(* CODESYS project cognex_insight.library
   DefaultNamespace: KOSTAL.AF2024.Drivers.Camera.Cognex_InSight
   DocFormat: reStructuredText
   Description: Provides communication via TcpIp or Ethernet/IP to Cognex InSight cameras.
   Author: Frank Dümpelmann, Martí Puig (F2R Automation)
   Title: KOSTAL.AF2024.Drivers.Camera.Cognex_InSight
   Version: 3.0.0.0
   Company: KOSTAL GmbH & Co.KG
   Placeholder: KOSTAL.AF2024.Drivers.Camera.Cognex_InSight

Project tree, tasks and I/O mapping:
  libraries: KOSTAL.AF2024.Core.ListOf, 1.0.0.0 (KOSTAL GmbH & Co.KG); KOSTAL.AF2024.Core.Process, 1.1.0.0 (KOSTAL GmbH & Co.KG); KOSTAL.AF2024.Core.Settings, 1.0.0.0 (KOSTAL GmbH & Co.KG); KOSTAL.AF2024.Core.StringTools, 1.0.0.0 (KOSTAL GmbH & Co.KG); KOSTAL.AF2024.Core.System, 1.0.0.0 (KOSTAL GmbH & Co.KG); KOSTAL.AF2024.Drivers.Camera.I_Camera, 2.0.0.0 (KOSTAL GmbH & Co.KG); Tc2_Standard, 3.4.5.0 (Beckhoff Automation GmbH); Tc2_System, 3.9.1.0 (Beckhoff Automation GmbH); Tc2_TcpIp, 3.4.2.0 (Beckhoff Automation GmbH); Tc2_Utilities, 3.9.2.0 (Beckhoff Automation GmbH)
  EthernetIP/
    DUT/
      Result/
        interface I_T_Result_Base: Clear, ResultArray
      data type _E_THIS_EIP
      data type _T_InspectionResult
      data type ST_IN_EIP
      data type ST_OUT_EIP
    function block FB_InSight_EIP [ST]: _a0_StepFail, _a0_StepInit, _a1_finish, _a1_idle, _a2_callTrigger, _a2_changeProgNum, _a2_inspection_Result, _connectControl, _FBmain, _resetfault, Ex_SetProgramNumber, Ex_Trigger, Ex_Trigger_ProgramNumber, FaultReset, LinkResult, Fault, ProgNo, ResultPass, State, FBmain
    interface I_InSight_EIP: Fault
  Project Information/
    function F_GetCompany [ST]
    function F_GetTitle [ST]
    function F_GetVersion [ST]
  TcpIp/
    DUT/
      Info/
        interface I_T_Info_TcpIp: ApplicationVersion, CopyTo, DateOfBuild, MacAddress, MonitorVersion, SerialNumber
        interface I_T_Info_TcpIp_CopyFrom: CopyFrom
        interface I_T_Info_TcpIp_Owner: ApplicationVersion, Clear, CopyFrom, DateOfBuild, MacAddress, MonitorVersion, SerialNumber
        function block T_Info_TcpIp [ST]: ApplicationVersion, Clear, CopyFrom, CopyTo, DateOfBuild, MacAddress, MonitorVersion, SerialNumber
      Internal/
        data type _E_PrgType_TcpIp
        data type _E_THIS_TcpIp
      data type E_BuilderVersion_TcpIp
      data type E_Command_TcpIp
      data type E_ProgLocation_TcpIp
    function block FB_InSight_Explorer_TcpIp [ST]: FB_init, _c1_Receive, _c1_Send, _c1_Socket, _connectionInit, _catchMacId, _catchPrgId, _catchPrgName, _foundEtx, _isCommandAccept, _isPasswordRequest, _isUserAccrepted, _isUserRequest, _isWelcome, _SplitData, _getCommand, _a3_GetData, _a3_GetData_DS, _a3_GetData_ETH, _a0_stepFail, _a0_stepInit, _a1_failure, _a1_Finish, _a1_Idle, _a2_Login, _a3_GetInfo, _a3_GetPrgId, _a3_GetPrgName, _a3_SetOffline, _a3_SetOnline, _a3_SetReqPrgById, _a3_SetReqPrgByName, _a3_Trigger, _FBmain, Ex_GetInfo, Ex_GetProgamNumber, Ex_GetProgramName, Ex_SetProgramName, Ex_SetProgramNumber, Ex_Trigger, Ex_Trigger_ProgName, Ex_Trigger_ProgramNumber, CommandPort, CommandTimeOut, IP, Data, DigitalSignalRuntime, DisableComplexResult, Info, ProgLocation, ResultPass, State, FBmain
    function block FB_InSight_VisionSuite_TcpIp [ST]: _catchMacId, _getCommand, SheetName
    interface I_InSight_TcpIp: Ex_GetInfo, Ex_GetProgamNumber, Ex_GetProgramName, Ex_SetProgramName, Ex_Trigger_ProgName, CommandPort, CommandTimeOut, IP, Data, DigitalSignalRuntime, DisableComplexResult, Info, ProgLocation
  Version/
    global variables Global_Version
*)

// EthernetIP/DUT/_E_THIS_EIP
{attribute 'qualified_only'}
{attribute 'strict'}
TYPE INTERNAL _E_THIS_EIP :
(
	idle	:= 0,
	trig,			
	trigPrgNum,
	chgprgnum	
) UINT;
END_TYPE

// EthernetIP/DUT/_T_InspectionResult
TYPE INTERNAL _T_InspectionResult : ARRAY[1..480] OF BYTE; END_TYPE

// EthernetIP/DUT/ST_IN_EIP
{attribute 'pack_mode' := '0'} 
TYPE ST_IN_EIP :
	STRUCT	
		TriggerReady 					: BIT;		//0.0
		TriggerACK						: BIT;		//0.1
		noName_0_0						: BIT;		//0.2
		MissedAcq							: BIT;		//0.3
		OfflineReason_1				: BIT;		//0.4		
		OfflineReason_2				: BIT;		//0.5
		OfflineReason_3				: BIT;		//0.6
		Online								: BIT;		//0.7
		SystemBusy						: BIT;		//1.0
		InspectionCompleted		: BIT;      //1.1
		ResultsBufferOverrun	: BIT;      //1.2
		ResultsValid					: BIT;      //1.3
		CommandExecuting			: BIT;      //1.4
		CommandComplete				: BIT;      //1.5
		CommandFailed					: BIT;      //1.6
		Error									: BIT;      //1.7
		SetUserDataAck				: BIT;		//2.0
		noName_1_0						: BIT;      //2.1
		noName_1_1						: BIT;      //2.2
		ExposureComplete			: BIT;      //2.3
		JobPass								: BIT;      //2.4
		TestRunReady					: BIT;      //2.5
		noName_2_0						: BIT;      //2.6
		noName_2_1						: BIT;      //2.7
		SoftEventACK_0				: BIT;		//3.0
		SoftEventACK_1				: BIT;      //3.1
		SoftEventACK_2				: BIT;      //3.2
		SoftEventACK_3				: BIT;      //3.3
		SoftEventACK_4				: BIT;      //3.4
		SoftEventACK_5				: BIT;      //3.5
		SoftEventACK_6				: BIT;      //3.6
		SoftEventACK_7				: BIT;      //3.7
		ErrorCode							: INT;
		noName_3_0						: BYTE;
		noName_3_1						: BYTE;
		CurrentJobID					: UINT;		
		AcquisitionID					: UINT;
		IspectionID						: UINT;
		InspectionResultCode	: INT;
		InspectionResult			: _T_InspectionResult;
	END_STRUCT
END_TYPE

// EthernetIP/DUT/ST_OUT_EIP
{attribute 'pack_mode' := '0'} 
TYPE ST_OUT_EIP :
	STRUCT
		TriggerEnable					: BIT; 		//0.0								
		Trigger								: BIT; 	    //0.1
		BufferResultsEnable		: BIT; 	    //0.2
		InspectionResultsACK	: BIT; 	    //0.3
		ExecuteCommand				: BIT; 	    //0.4
		noName_0_0						: BIT; 	    //0.5
		noName_0_1						: BIT; 	    //0.6
		SetOffline						: BIT; 	    //0.7
		noName_1							: BYTE;		//1
		SetUserData						: BIT; 		//2.0
		noName_2_0						: BIT; 	    //2.1
		ClearError						: BIT; 	    //2.2
		ClearExposureComplete	: BIT; 	    //2.3
		noName_3_0						: BIT; 	    //2.4
		noName_3_1						: BIT;      //2.5
		noName_3_2						: BIT; 	    //2.6
		noName_3_3						: BIT;      //2.7
		SoftEvent_0						: BIT; 		//3.0
		SoftEvent_1						: BIT;      //3.1
		SoftEvent_2						: BIT;      //3.2
		SoftEvent_3						: BIT;      //3.3
		SoftEvent_4						: BIT;      //3.4
		SoftEvent_5						: BIT;      //3.5
		SoftEvent_6						: BIT;      //3.6
		SoftEvent_7						: BIT;      //3.7
		CommandID							: UINT;	
		noName_4_0						: BYTE; 	
		noName_4_1						: BYTE; 	
		UserData							: _T_InspectionResult;// ARRAY[0..487] OF BYTE; 
	END_STRUCT
END_TYPE

// TcpIp/DUT/Internal/_E_PrgType_TcpIp
{attribute 'qualified_only'}
{attribute 'strict'}
TYPE INTERNAL _E_PrgType_TcpIp :
(
	Number := 0,
	Name
) UINT;
END_TYPE

// TcpIp/DUT/Internal/_E_THIS_TcpIp
{attribute 'qualified_only'}
{attribute 'strict'}
TYPE INTERNAL _E_THIS_TcpIp :
(
	Idle := 0,
	GetInfo,

	Trigger,
	TriggerPrgNo,
	TriggerPrgName,

	SetOnline,
	GetOnline,

	SetProgramId,
	GetProgramId,

	SetProgramName,
	GetProgramName,

	ReadVersion,
	ReadOperationMode
) UINT;
END_TYPE

// TcpIp/DUT/E_BuilderVersion_TcpIp
{attribute 'qualified_only'}
{attribute 'strict'}
TYPE E_BuilderVersion_TcpIp :
(
	InSightExplorer 	:= 0,
	InSigtVisionSuite	:= 1
);
END_TYPE

// TcpIp/DUT/E_Command_TcpIp
{attribute 'qualified_only'}
{attribute 'strict'}
TYPE E_Command_TcpIp :
(
	GetInfo := 0,
	UserName,
	Password,
	SetOnline,
	SetOffline,
	GetOnline,
	GetPrgId,
	SetPrgId,
	GetPrgName,
	SetPrgName,
	Trigger,
	GetFormatstring
);
END_TYPE

// TcpIp/DUT/E_ProgLocation_TcpIp
{attribute 'qualified_only'}
{attribute 'strict'}
TYPE E_ProgLocation_TcpIp :
(
	None := 0,
	FlashMemory,
	RamDisk,
	SD_Card
);
END_TYPE

// Version/Global_Version
{attribute 'TcGenerated'}
{attribute 'no-analysis'}
{attribute 'linkalways'}
// This function has been automatically generated from the project information.
VAR_GLOBAL CONSTANT
	{attribute 'const_non_replaced'}
	stLibVersion_KOSTAL_AF2024_Drivers_Camera_Cognex_InSight : ST_LibVersion := (iMajor := 3, iMinor := 0, iBuild := 0, iRevision := 0, nFlags := 0, sVersion := '3.0.0.0');
END_VAR

// EthernetIP/DUT/Result/I_T_Result_Base
INTERFACE PUBLIC I_T_Result_Base EXTENDS KOSTAL_AF2024_Core_System.I_Interface

METHOD PUBLIC Clear
VAR

END_VAR
END_METHOD

PROPERTY PUBLIC ResultArray : REFERENCE TO _T_InspectionResult
GET
END_GET
END_PROPERTY

END_INTERFACE

// EthernetIP/FB_InSight_EIP
FUNCTION_BLOCK FB_InSight_EIP IMPLEMENTS I_InSight_EIP//, _I_T_Result

VAR
	{region 'EthernetIP Communications'}
		ECatState			AT %I*	: UINT;	//link to EtherCat State from {Device x (ECAT EIP Scanner (EL6652))}.Inputs.State
		InSightState	AT %I*	: UINT;	//link to {InSight 2000 Series}.Inputs.State
	
		InSight_IN 	AT %I*	: ST_IN_EIP; //link with Continious mode ATTENTION be sure, that the Array-Nodes are collapsed
		InSight_OUT AT %Q*	: ST_OUT_EIP; //link with Continious mode ATTENTION be sure, that the Array-Nodes are collapsed
															
//		InSight_IN	: POINTER TO ST_IN_EIP;
//		InSight_OUT	: POINTER TO ST_OUT_EIP;
	{endregion}
                            	                     	
	_step	: KOSTAL_AF2024_Core_Process.FB_processStep_Flow;	//Use the “_Flow” step to save runtime. 

	_THIS_CALLED			: _E_THIS_EIP;
	_THIS_IN_PROCESS	: _E_THIS_EIP;

	_state	: KOSTAL_AF2024_Core_Process.T_plcState;
	
	{region 'Functionality'}
		//Inputs 
		_Reset	: BOOL;
		_prgNum	: UINT;
															
		//Outputs               	
		_InspectionOK				: BOOL;
		//_InspectionNOK			: BOOL;
		//_refResult	: REFERENCE TO _T_InspectionResult;
		_Iresult	: I_T_Result_Base;	 
 
	{endregion}

	{region 'Static'}
		TON_Change_Job : Tc2_Standard.TON;
	{endregion}
		 

	
		 
	
END_VAR

VAR CONSTANT
	_ADDRESS_Idle						: INT:= 0;
	_ADDRESS_TriggerPrgNum	: INT:= 100;	//Job ID
	_ADDRESS_SetPrgNum			: INT:= 200;	//Job ID
END_VAR

METHOD PROTECTED _a0_StepFail
VAR_INPUT
END_VAR

_state.clear();
_state.fail:= TRUE;
_state.description:= Tc2_Standard.WCONCAT(INT_TO_WSTRING(_step.actual), ". Step does not exist");
END_METHOD

METHOD PROTECTED _a0_StepInit
VAR_INPUT
END_VAR

IF (_THIS_CALLED <> _THIS_IN_PROCESS) AND_THEN (_step.actual <> _ADDRESS_Idle) THEN	_step.init();	END_IF
END_METHOD

METHOD PROTECTED _a1_finish 
VAR_INPUT
END_VAR

_state.clear();

_state.finish := TRUE;
_state.pass:= TRUE;
END_METHOD

METHOD PROTECTED _a1_idle

//Idle process - Clear information from other processes
IF _step.toggle THEN

	InSight_OUT.Trigger								:= FALSE;
	InSight_OUT.TriggerEnable					:= FALSE;
	InSight_OUT.InspectionResultsACK := FALSE;

END_IF


_state.clear();

IF _THIS_CALLED = _E_THIS_EIP.idle THEN

	_THIS_IN_PROCESS:= _THIS_CALLED;

	_state.ready := TRUE;

	
ELSIF _THIS_CALLED = _E_THIS_EIP.chgprgnum THEN

	_THIS_IN_PROCESS:= _THIS_CALLED;

	_state.busy := TRUE;

	_step.set(_ADDRESS_SetPrgNum);
	
	
ELSIF _THIS_CALLED = _E_THIS_EIP.trigPrgNum THEN

	_THIS_IN_PROCESS:= _THIS_CALLED;

	_state.busy := TRUE;

	_InspectionOK:= FALSE;
	
	_step.set(_ADDRESS_TriggerPrgNum);

	
ELSIF _THIS_CALLED = _E_THIS_EIP.trig THEN

	_THIS_IN_PROCESS:= _THIS_CALLED;

	_state.busy := TRUE;

	_InspectionOK:= FALSE;

	_step.set(_ADDRESS_TriggerPrgNum);
	
ELSE

	_THIS_IN_PROCESS:= _E_THIS_EIP.idle;

	_state.finish	:= TRUE;
	_state.fail		:= TRUE;
	_state.description:= 	"Process with this enumeration does not exist!"; 

END_IF
END_METHOD

METHOD PROTECTED _a2_callTrigger
VAR_INPUT
END_VAR

VAR_INST	
	_SubStep		: KOSTAL_AF2024_Core_Process.FB_processStep_Flow;
	_PF_InspectionCompleted	:BOOL;
END_VAR

IF _step.toggle THEN	
	_subStep.init();
	IF _Iresult <> 0 THEN
		_Iresult.Clear();
END_IF	
END_IF

_state.description:= "Method _a2_callTrigger() is running ...";

InSight_OUT.InspectionResultsACK := FALSE;

_subStep.Header();

IF _SubStep.isActive(0) THEN IF InSight_IN.ResultsValid THEN InSight_OUT.InspectionResultsACK := TRUE; ELSE _SubStep.INC(); END_IF END_IF
	
IF _SubStep.isActive(1) THEN IF NOT  InSight_IN.ResultsValid THEN InSight_OUT.TriggerEnable := TRUE ; InSight_OUT.InspectionResultsACK := FALSE; _SubStep.INC(); END_IF END_IF

IF _SubStep.isActive(2) THEN IF  InSight_IN.TriggerReady (*AND NOT _pIN^.InspectionCompleted*) THEN InSight_OUT.Trigger:= TRUE; _SubStep.INC(); END_IF END_IF

IF _SubStep.isActive(3) THEN IF InSight_IN.InspectionCompleted <> _PF_InspectionCompleted THEN InSight_OUT.Trigger := FALSE; _step.INC(); END_IF END_IF

_PF_InspectionCompleted := InSight_IN.InspectionCompleted;
END_METHOD

METHOD PROTECTED _a2_changeProgNum
VAR_INPUT
END_VAR
IF _step.toggle THEN	;	END_IF

_state.description:= "Method _a2_changeProgNum() is running ...";

IF InSight_IN.CurrentJobID > 0 AND InSight_IN.CurrentJobID = _prgNum THEN
	
	InSight_OUT.SetOffline := FALSE;
	TON_Change_Job(IN:= FALSE);

	_step.INC();

ELSE

	InSight_OUT.CommandID := _prgNum;
	InSight_OUT.SetOffline := TRUE;

	IF  NOT InSight_IN.Online AND InSight_IN.OfflineReason_1 THEN
		//TON_Change_Job.PT := T#100MS;
		//TON_Change_Job.IN := TRUE;
		TON_Change_Job(IN:= TRUE, PT:= T#100MS, Q=> , ET=> );
	END_IF

END_IF

InSight_OUT.ExecuteCommand := TON_Change_Job.Q;
END_METHOD

METHOD PROTECTED _a2_inspection_Result
VAR_INPUT
END_VAR

IF _step.toggle THEN	;	END_IF

_state.description:= "Method _a2_inspection_Result() is running ...";

InSight_OUT.TriggerEnable 	:= FALSE ;
_InspectionOK  				:= FALSE;


IF _Iresult <> 0 AND_THEN __ISVALIDREF(_Iresult.ResultArray) THEN
	_Iresult.ResultArray := InSight_IN.InspectionResult;
END_IF


_InspectionOK := InSight_IN.InspectionResult[1] = 1;

_step.INC();
END_METHOD

METHOD PROTECTED _connectControl : BOOL
VAR_INPUT
END_VAR

 
IF ECatState <> 0  THEN

	_connectControl:= FALSE;

	_state.clear();
	_state.fail:= TRUE;
	_state.description:= Tc2_Standard.WCONCAT(UINT_TO_WSTRING(ECatState), ";Error from EtherCAT (EIP-Scanner)");


	_step.init();

ELSIF InSightState <> 0 THEN

	_connectControl:= FALSE;

	_state.clear();
	_state.fail:= TRUE;
	_state.description:= Tc2_Standard.WCONCAT(UINT_TO_WSTRING(InSightState), ";Error from Ethernet IP Connection");

	_step.init();

ELSE
	
	_connectControl:= TRUE;

END_IF
END_METHOD

METHOD PROTECTED _FBmain
VAR_INPUT
END_VAR
// is set duriing FB_Init() method
//_pIN:= ADR(InSight2000_IN[2]);
//_pOUT:= ADR(InSight2000_OUT[2]);


IF NOT _connectControl() THEN RETURN;	END_IF

_a0_StepInit();

_step.Header();

IF _step.isActive(_ADDRESS_Idle) THEN _a1_idle();	END_IF


//Trigger and TriggerPrgNum uses the same steps
IF _step.isActive(_ADDRESS_TriggerPrgNum)			THEN _step.INC();							END_IF
IF _step.isActive(_ADDRESS_TriggerPrgNum + 1)	THEN _a2_changeProgNum();			END_IF
IF _step.isActive(_ADDRESS_TriggerPrgNum + 2)	THEN _a2_callTrigger();				END_IF
IF _step.isActive(_ADDRESS_TriggerPrgNum + 3)	THEN _a2_inspection_Result();	END_IF
IF _step.isActive(_ADDRESS_TriggerPrgNum + 4)	THEN _a1_finish();						END_IF


IF _step.isActive(_ADDRESS_SetPrgNum)			THEN _step.INC();					END_IF
IF _step.isActive(_ADDRESS_SetPrgNum + 1)	THEN _a2_changeProgNum();	END_IF
IF _step.isActive(_ADDRESS_SetPrgNum + 2)	THEN _a1_finish();				END_IF


IF _step.NotFound() THEN _a0_StepFail();	END_IF

_resetfault();
END_METHOD

METHOD PROTECTED _resetfault
VAR_INPUT
END_VAR

IF _Reset AND InSight_IN.Error THEN	InSight_OUT.ClearError := TRUE;
ELSE														InSight_OUT.ClearError := FALSE;
END_IF

_Reset:= FALSE;
END_METHOD

METHOD PUBLIC Ex_SetProgramNumber : BOOL;
VAR_INPUT
	ProgramNumber : UINT;
END_VAR
IF _THIS_CALLED = _E_THIS_EIP.idle THEN //Another process is running: don't start this process!

	_prgNum := ProgramNumber;
	
	_THIS_CALLED := _E_THIS_EIP.chgprgnum;
	
	_FBmain();	//Call sequence via _FBmain
	
	Ex_SetProgramNumber := _THIS_CALLED = _THIS_IN_PROCESS;	//Return true when process was started
	
END_IF
END_METHOD

METHOD Ex_Trigger : BOOL

IF _THIS_CALLED = _E_THIS_EIP.idle THEN //Another process is running: don't start this process!

	_THIS_CALLED := _E_THIS_EIP.trig;
	
	_FBmain();	//Call sequence via _FBmain
	
	Ex_Trigger := _THIS_CALLED = _THIS_IN_PROCESS;	//Return true when process was started

END_IF
END_METHOD

METHOD PUBLIC Ex_Trigger_ProgramNumber : BOOL;
VAR_INPUT
	ProgramNumber : UINT;
END_VAR
IF _THIS_CALLED = _E_THIS_EIP.idle THEN //Another process is running: don't start this process!

	IF ProgramNumber <> 0 THEN	_prgNum := ProgramNumber;	END_IF
	
	_THIS_CALLED := _E_THIS_EIP.trigPrgNum;
	
	_FBmain();	//Call sequence via _FBmain
	
	Ex_Trigger_ProgramNumber := _THIS_CALLED = _THIS_IN_PROCESS;	//Return true when process was started

END_IF
END_METHOD

METHOD PUBLIC FaultReset

_Reset := TRUE;
END_METHOD

METHOD PUBLIC LinkResult
VAR_INPUT
	result 	: I_T_Result_Base;
END_VAR
IF result <> 0 THEN
 _Iresult := result; 
END_IF;
END_METHOD

PROPERTY Fault : bool
GET
Fault := InSight_IN.Error;
END_GET
END_PROPERTY

PROPERTY ProgNo : UINT
GET

ProgNo:=  InSight_IN.CurrentJobID;;
END_GET
END_PROPERTY

PROPERTY ResultPass : BOOL
GET

ResultPass:= _InspectionOK;
END_GET
END_PROPERTY

PROPERTY State : KOSTAL_AF2024_Core_Process.I_T_plcState
GET
State := _state;
END_GET
END_PROPERTY

METHOD FBmain
VAR_INPUT
END_VAR

VAR

END_VAR

IF _THIS_CALLED = _E_THIS_EIP.idle THEN
	_FBmain();
END_IF
_THIS_CALLED:= _E_THIS_EIP.idle;
END_METHOD

END_FUNCTION_BLOCK

// EthernetIP/I_InSight_EIP
INTERFACE I_InSight_EIP EXTENDS KOSTAL_AF2024_Drivers_Camera_I_Camera.I_Camera

PROPERTY Fault : bool
GET
END_GET
END_PROPERTY

END_INTERFACE

// Project Information/F_GetCompany
// This function has been automatically generated from the project information.
{attribute 'signature_flag' := '1073741824'}
{attribute 'TcGenerated'}
{attribute 'no-analysis'}
FUNCTION F_GetCompany : WSTRING
VAR_INPUT
	
END_VAR

F_GetCompany := "KOSTAL GmbH & Co.KG";

END_FUNCTION

// Project Information/F_GetTitle
// This function has been automatically generated from the project information.
{attribute 'signature_flag' := '1073741824'}
{attribute 'TcGenerated'}
{attribute 'no-analysis'}
FUNCTION F_GetTitle : WSTRING
VAR_INPUT
	
END_VAR

F_GetTitle := "KOSTAL.AF2024.Drivers.Camera.Cognex_InSight";

END_FUNCTION

// Project Information/F_GetVersion
// This function has been automatically generated from the project information.
{attribute 'signature_flag' := '1073741824'}
{attribute 'TcGenerated'}
{attribute 'no-analysis'}
FUNCTION F_GetVersion : ST_LibVersion
VAR_INPUT
	
END_VAR

F_GetVersion.iMajor := 3;
F_GetVersion.iMinor := 0;
F_GetVersion.iBuild := 0;
F_GetVersion.iRevision := 0;
F_GetVersion.sVersion := '3.0.0.0';
F_GetVersion.nFlags := 0;

END_FUNCTION

// TcpIp/DUT/Info/I_T_Info_TcpIp
INTERFACE I_T_Info_TcpIp EXTENDS KOSTAL_AF2024_Core_System.I_Interface

PROPERTY PUBLIC ApplicationVersion : KOSTAL_AF2024_Core_Settings.T_MaxString_UTF8
GET
END_GET
END_PROPERTY

METHOD PUBLIC CopyTo : BOOL
VAR_INPUT
	IN	: I_T_Info_TcpIp_CopyFrom;
END_VAR
END_METHOD

PROPERTY PUBLIC DateOfBuild : KOSTAL_AF2024_Core_Settings.T_MaxString_UTF8
GET
END_GET
END_PROPERTY

PROPERTY PUBLIC MacAddress : KOSTAL_AF2024_Core_Settings.T_MaxString_UTF8
GET
END_GET
END_PROPERTY

PROPERTY PUBLIC MonitorVersion : KOSTAL_AF2024_Core_Settings.T_MaxString_UTF8
GET
END_GET
END_PROPERTY

PROPERTY PUBLIC SerialNumber : KOSTAL_AF2024_Core_Settings.T_MaxString_UTF8
GET
END_GET
END_PROPERTY

END_INTERFACE

// TcpIp/DUT/Info/I_T_Info_TcpIp_CopyFrom
INTERFACE I_T_Info_TcpIp_CopyFrom EXTENDS KOSTAL_AF2024_Core_System.I_Interface

METHOD PUBLIC CopyFrom : BOOL
VAR_INPUT
	IN	: KOSTAL_AF2024_Core_System.I_Interface;
END_VAR
END_METHOD

END_INTERFACE

// TcpIp/DUT/Info/I_T_Info_TcpIp_Owner
INTERFACE I_T_Info_TcpIp_Owner EXTENDS I_T_Info_TcpIp

PROPERTY PUBLIC ApplicationVersion : KOSTAL_AF2024_Core_Settings.T_MaxString_UTF8
SET
END_SET
END_PROPERTY

METHOD PUBLIC Clear
VAR_INPUT
END_VAR
END_METHOD

METHOD PUBLIC CopyFrom : BOOL
VAR_INPUT
	IN	: KOSTAL_AF2024_Core_System.I_Interface;
END_VAR
END_METHOD

PROPERTY PUBLIC DateOfBuild : KOSTAL_AF2024_Core_Settings.T_MaxString_UTF8
SET
END_SET
END_PROPERTY

PROPERTY PUBLIC MacAddress : KOSTAL_AF2024_Core_Settings.T_MaxString_UTF8
SET
END_SET
END_PROPERTY

PROPERTY PUBLIC MonitorVersion : KOSTAL_AF2024_Core_Settings.T_MaxString_UTF8
SET
END_SET
END_PROPERTY

PROPERTY PUBLIC SerialNumber : KOSTAL_AF2024_Core_Settings.T_MaxString_UTF8
SET
END_SET
END_PROPERTY

END_INTERFACE

// TcpIp/DUT/Info/T_Info_TcpIp
FUNCTION_BLOCK PUBLIC T_Info_TcpIp IMPLEMENTS I_T_Info_TcpIp, I_T_Info_TcpIp_Owner, I_T_Info_TcpIp_CopyFrom

VAR
	_SerialNumber				: KOSTAL_AF2024_Core_Settings.T_MaxString_UTF8;
	_ApplicationVersion	: KOSTAL_AF2024_Core_Settings.T_MaxString_UTF8;
	_MonitorVersion			: KOSTAL_AF2024_Core_Settings.T_MaxString_UTF8;
	_MacAddress					: KOSTAL_AF2024_Core_Settings.T_MaxString_UTF8;
	_DateOfBuild				: KOSTAL_AF2024_Core_Settings.T_MaxString_UTF8;
END_VAR

PROPERTY PUBLIC ApplicationVersion : KOSTAL_AF2024_Core_Settings.T_MaxString_UTF8
GET

ApplicationVersion:= _ApplicationVersion;
END_GET
SET

_ApplicationVersion:= ApplicationVersion;
END_SET
END_PROPERTY

METHOD PUBLIC Clear

_SerialNumber				:= '';
_ApplicationVersion	:= '';
_MonitorVersion			:= '';
_MacAddress					:= '';
_DateOfBuild				:= '';
END_METHOD

METHOD PUBLIC CopyFrom : BOOL
VAR_INPUT
	IN	: KOSTAL_AF2024_Core_System.I_Interface;
END_VAR

VAR
	_obj	: I_T_Info_TcpIp;
END_VAR

IF (IN = 0) OR_ELSE NOT __QUERYINTERFACE(IN, _obj) OR_ELSE (_obj = 0) THEN RETURN;	END_IF

_SerialNumber				:= _obj.SerialNumber;
_ApplicationVersion	:= _obj.ApplicationVersion;
_MonitorVersion			:= _obj.MonitorVersion;
_MacAddress					:= _obj.MacAddress;
_DateOfBuild				:= _obj.DateOfBuild;

CopyFrom:= TRUE;
END_METHOD

METHOD PUBLIC CopyTo : BOOL
VAR_INPUT
	IN	: I_T_Info_TcpIp_CopyFrom;
END_VAR

VAR
	_obj	: I_T_Info_TcpIp_CopyFrom;
END_VAR

IF (IN = 0) OR_ELSE NOT __QUERYINTERFACE(IN, _obj) OR_ELSE (_obj = 0) THEN RETURN;	END_IF

CopyTo:= IN.CopyFrom(THIS^);
END_METHOD

PROPERTY PUBLIC DateOfBuild : KOSTAL_AF2024_Core_Settings.T_MaxString_UTF8
GET

DateOfBuild:= _DateOfBuild;
END_GET
SET

_DateOfBuild:= DateOfBuild;
END_SET
END_PROPERTY

PROPERTY PUBLIC MacAddress : KOSTAL_AF2024_Core_Settings.T_MaxString_UTF8
GET

MacAddress:= _MacAddress;
END_GET
SET

_MacAddress:= MacAddress;
END_SET
END_PROPERTY

PROPERTY PUBLIC MonitorVersion : KOSTAL_AF2024_Core_Settings.T_MaxString_UTF8
GET

MonitorVersion:= _MonitorVersion;
END_GET
SET

_MonitorVersion:= MonitorVersion;
END_SET
END_PROPERTY

PROPERTY PUBLIC SerialNumber : KOSTAL_AF2024_Core_Settings.T_MaxString_UTF8
GET

SerialNumber:= _SerialNumber;
END_GET
SET

_SerialNumber:= SerialNumber;
END_SET
END_PROPERTY

END_FUNCTION_BLOCK

// TcpIp/FB_InSight_Explorer_TcpIp
FUNCTION_BLOCK PUBLIC FB_InSight_Explorer_TcpIp IMPLEMENTS I_InSight_TcpIp

VAR CONSTANT
		_CMD_PORT_DEFAULT		: UDINT:= 23;
		_DATA_PORT_DEFAULT	: UDINT:= 9004;

		_ETX								: STRING(2)		:= '$0D$0A';
		_JOB_EXTENSION 			: STRING(4):= '.job';

		_STORAGE_FLASH_MEMORY	: STRING:= '';
		_STORAGE_RAM_DISK			: STRING:= 'RAMDisk';
		_STORAGE_SD_CARD			: STRING:= 'SDCARD';
		
		_DEFAULT_TIMEOUT	: TIME:= T#5S;
END_VAR

VAR

	{region 'Connection'}
		_ServerAmsNetId	: Tc2_System.T_AmsNetID:= '';
		_IP							: Tc2_System.T_IPv4Addr;
		_CmdPort				: UDINT:= _CMD_PORT_DEFAULT;
		_DataPort				: UDINT:= _DATA_PORT_DEFAULT;
	{endregion}

	{region 'Command'}
		_cmdSocket							: Tc2_TcpIp.FB_ClientServerConnection;
		_CmdExecutedSocketState	:	Tc2_TcpIp.E_SocketConnectionState;
		_cmdSend								: Tc2_TcpIp.FB_SocketSend;
		_cmdReceive							: Tc2_TcpIp.FB_SocketReceive;

		_cmdTimeOut			: TIME	:= T#5S;	//default T#5S
		_cmdSocketTimer	: TON;	//TON

		_cmdReceivedPartly	: KOSTAL_AF2024_Core_Settings.T_MaxString_UTF8;
		_cmdReceivedString	: KOSTAL_AF2024_Core_Settings.T_MaxString_UTF8;
		_cmdResponse				: KOSTAL_AF2024_Core_Settings.T_MaxString_UTF8;

		_Cmd		: KOSTAL_AF2024_Core_Settings.T_MaxString_UTF8;
	{endregion}

	{region 'Data'}
		_dataResponse				: KOSTAL_AF2024_Core_Settings.T_MaxString_UTF8;
		_Data			: KOSTAL_AF2024_Core_ListOf.FB_ListOfString_UTF8;	
	{endregion}
	
	_Info	: T_Info_TcpIp;

	_PrgNum			: UINT:= 1;	//Job ID - default 1
	_PrgNumResp	: UINT;	//Job ID - last responsed program number

	_PrgName			: KOSTAL_AF2024_Core_Settings.T_MaxString_UTF8;	//Job File Name 
	_PrgNameResp	: KOSTAL_AF2024_Core_Settings.T_MaxString_UTF8;	//Job File Name - last responsed program name
	
	_PrgLocation 			: E_ProgLocation_TcpIp:= E_ProgLocation_TcpIp.FlashMemory;	//define the location of stored programs - default
	_PrgLocationResp	: E_ProgLocation_TcpIp:= E_ProgLocation_TcpIp.None;			//last response of file on storage 
	
	_Step		: KOSTAL_AF2024_Core_Process.FB_processStep_Flow;
	_State	:	KOSTAL_AF2024_Core_Process.T_plcState;

	_THIS_CALLED			: _E_THIS_TcpIp;
	_THIS_IN_PROCESS	: _E_THIS_TcpIp;

	_Init			: BOOL:= TRUE;

	{region 'Digital Signal'}
		_DisableComplexResult		: BOOL;	//Use this parameter to link the result of the camera inspection only to the digital PASS channel.
		_DigitalSignalRuntime		: TIME:= T#150MS;	//Waiting time before the digital signal is analyzed.
		_DigitalSignalRuntimer	: TON;
		_DigitalSignal	AT %I*	:	BOOL;	//Digital PASS Input signal
	{endregion}

END_VAR

VAR CONSTANT
	_ADDRESS_GetInfo				: INT:= 100;

	_ADDRESS_Trigger				: INT:= 200;	//no program check
	_ADDRESS_TriggerPrgNum	: INT:= 300;	//Job ID
	_ADDRESS_TriggerPrgName	: INT:= 400;	//Job File Name

	_ADDRESS_SetPrgNum			: INT:= 500;	//Job ID
	_ADDRESS_GetPrgNum			: INT:= 600;	//Job ID

	_ADDRESS_SetPrgName			: INT:= 700;	//Job name
	_ADDRESS_GetPrgName			: INT:= 800;	//Job name
END_VAR

METHOD FB_init : BOOL
VAR_INPUT
	bInitRetains : BOOL; // if TRUE, the retain variables are initialized (warm start / cold start)
	bInCopyCode : BOOL;  // if TRUE, the instance afterwards gets moved into the copy code (online change)

	ServerAmsNetId	: Tc2_System.T_AmsNetID;	//AmsNetId of TcpIp-Server Provider - default local > ''

	IP					: Tc2_System.T_IPv4Addr;	//IP Address of camera system
	CommandPort	: UDINT;	//Entry 0 > default port will used
	DisableComplexResult	: BOOL;	//Use this parameter to link the result of the camera inspection only to the digital PASS channel.
END_VAR
IF IP <> '' 									THEN _IP:= IP;													END_IF 
IF ServerAmsNetId <> ''				THEN	_serverAmsNetId:= serverAmsNetId;	END_IF
IF CommandPort		<> UDINT#0	THEN	_CmdPort:= CommandPort;						END_IF

_DisableComplexResult:= DisableComplexResult;
END_METHOD

METHOD PROTECTED _c1_Receive : BOOL
VAR_INPUT
	Enable	:  BOOL;
	Toggle	: BOOL;
END_VAR
VAR_INST
	_onceReceived	: BOOL;
	_zeroRecs			: UINT;
END_VAR
IF Toggle THEN

	_cmdReceivedString:= '';
	_cmdReceivedPartly:= '';
	_cmdResponse			:= '';

	_onceReceived	:= FALSE;
	_zeroRecs			:= 0;
	
	_cmdReceive
	(
		bExecute:= FALSE,
		sSrvNetId	:= _serverAmsNetId,
		hSocket		:= _cmdSocket.hSocket,
		cbLen			:= SIZEOF(_cmdReceivedPartly) - 1,
		pDest			:= ADR(_cmdReceivedPartly),
		tTimeout	:= _cmdTimeOut
	);

END_IF


IF NOT Enable THEN	_cmdReceive(bExecute:= FALSE, hSocket:= _cmdSocket.hSocket);

ELSIF _c1_Socket(TRUE)	THEN

	_cmdReceive(bExecute:= TRUE, hSocket:= _cmdSocket.hSocket);

	IF _cmdReceive.bBusy THEN	

		_State.clear();
		_state.busy	:= TRUE;
		_state.description:= "camera is busy(command receive); wait ...";
			
	ELSIF _cmdReceive.bError THEN

		_State.clear();
		_state.description:= Tc2_Standard.WCONCAT("Error during command receive. Errorcode>", UDINT_TO_WSTRING(_cmdReceive.nErrId));
		_state.fail	:= TRUE;
		_state.finish:= TRUE;	

	ELSIF _cmdReceive.nRecBytes <> 0 THEN 

		_onceReceived:= TRUE;
		_zeroRecs:= 0;
		
		_cmdResponse:= _cmdReceivedString:= Tc2_Standard.CONCAT(STR1:= _cmdReceivedString, STR2:=  Tc2_Standard.LEFT(STR:= _cmdReceivedPartly, SIZE:= UDINT_TO_INT(_cmdReceive.nRecBytes)));
		_cmdReceivedPartly:= '';

		_cmdReceive(bExecute:= FALSE);
		
	ELSE	

		_zeroRecs:= _zeroRecs + 1;

		IF _onceReceived AND (_zeroRecs > 5) THEN	_c1_Receive:= TRUE;	ELSE	_cmdReceive(bExecute:= FALSE);	END_IF

	END_IF

END_IF
END_METHOD

METHOD PROTECTED _c1_Send : BOOL
VAR_INPUT
	Enable	:  BOOL;
	Toggle	: BOOL;
END_VAR

IF Toggle THEN 

	_cmdSend
	(
		bExecute:= FALSE,
		sSrvNetId	:= _serverAmsNetId,
		hSocket		:= _cmdSocket.hSocket,
		cbLen			:= TO_UDINT(Tc2_Standard.LEN(_Cmd)),
		pSrc			:= ADR(_Cmd),
		tTimeout	:= _cmdTimeOut
	); 

END_IF


IF NOT Enable THEN
	
	_c1_Send:= NOT _cmdSend.bBusy;

ELSIF _c1_Socket(TRUE)	THEN

	_cmdSend(bExecute:= TRUE, hSocket:= _cmdSocket.hSocket); 
	
	IF _cmdSend.bBusy THEN	
	
		_State.clear();
		_state.busy	:= TRUE;
		_state.description:= "Command Send is busy(Send ...)";
	
	ELSIF _cmdSend.bError THEN
	
		_State.clear();
		_State.description:= Tc2_Standard.WCONCAT("Error during command Send. Errorcode>", UDINT_TO_WSTRING(_cmdSend.nErrId));
		_State.fail	:= TRUE;
		_State.finish:= TRUE;	
	
	ELSE	_c1_Send:= TRUE;
	
	END_IF

END_IF
END_METHOD

METHOD PROTECTED _c1_Socket : BOOL
VAR_INPUT
	Enable	: BOOL;
END_VAR
	
_cmdSocket
(
	bEnable			:= Enable,
	sSrvNetID		:= _serverAmsNetId,
	nMode				:= Tc2_TcpIp.CONNECT_MODE_ENABLEDBG,
	sRemoteHost	:= _IP,
	nRemotePort	:= _CmdPort, 
	tReconnect	:= T#60S//_cmdTimeOut 
);

IF _cmdSocketTimer.Q THEN

	_State.clear();
	_State.description:= "command socket connection cannot be established - Timeout";
	_State.fail	:= TRUE;
	_State.finish:= TRUE;	

ELSIF NOT Enable THEN

	IF  _cmdSocket.bBusy THEN
		
		_State.clear();
		_state.busy	:= TRUE;
		_state.description:= "Command socket is busy(disconnecting ...)";

	ELSIF _cmdSocket.hSocket.handle <> 0 THEN	_cmdSocketTimer.IN:= TRUE;
		
		_State.clear();
		_state.busy	:= TRUE;
		_state.description:= "Command socket is busy(wait for handle clearance ...)";

	ELSE	_c1_Socket:= TRUE;
	END_IF


ELSE

	IF _cmdSocket.bBusy THEN	_cmdSocketTimer.IN:= TRUE;
	
		_State.clear();
		_state.busy	:= TRUE;
		_state.description:= "Command socket is busy(connect ...)";
	
	ELSIF _cmdSocket.bError THEN
	
		_State.clear();
		_State.description:= Tc2_Standard.WCONCAT("Error during command socket open. Errorcode>", UDINT_TO_WSTRING(_cmdSocket.nErrId));
		_State.fail	:= TRUE;
		_State.finish:= TRUE;	
	
	ELSIF _cmdsocket.hSocket.handle = 0 THEN
	
		_State.clear();
		_State.description:= "no Handle from command socket";
		_State.fail	:= TRUE;
		_State.finish:= TRUE;
	
	ELSE	_CmdExecutedSocketState:= _cmdSocket.eState;	_c1_Socket:= TRUE;
	
	END_IF
	
END_IF

_cmdSocketTimer(IN:= NOT _c1_Socket, PT:= _cmdTimeOut, Q=> , ET=> );
END_METHOD

METHOD PROTECTED _connectionInit

_c1_Send(FALSE, TRUE);
_c1_Receive(FALSE, TRUE);
_c1_Socket(FALSE);
_cmdSocketTimer(IN:= FALSE);

//_d1_Receive(FALSE, TRUE);
//_d1_ServerReceive(FALSE, TRUE);
//_d1_Socket(FALSE);
//_dataSocketTimer(IN:= FALSE);

//Tc2_TcpIp.F_CreateServerHnd(	'','',_DataPort, Tc2_TcpIp.LISTEN_MODE_CLOSEALL, FALSE, hServer:= _dataHServer);

//_dataServer
//(	hServer:= _dataHServer,
//	eMode:= Tc2_TcpIp.eACCEPT_ALL,
//	sRemoteHost:= '',
//	nRemotePort:= _DataPort,
//	bEnable:= FALSE,
//	tReconnect:= T#1S
//);

//Tc2_TcpIp.F_CreateServerHnd(	'','',_DataPort, Tc2_TcpIp.LISTEN_MODE_CLOSEALL, FALSE, hServer:= _dataHServer);
//_dataServer(bEnable:= FALSE, hServer:= _dataHServer);
END_METHOD

//cameras with InSigtExplorer sends MAC ID with '-'
METHOD PROTECTED _catchMacId : KOSTAL_AF2024_Core_Settings.T_MaxString_UTF8
VAR_INPUT
	IN	: KOSTAL_AF2024_Core_Settings.T_MaxString_UTF8;
END_VAR

//cameras with InSigtVisionSuite sends MAC ID with ':'

_catchMacId:= IN;
END_METHOD

METHOD PROTECTED _catchPrgId : BOOL

VAR_INPUT
	Toggle	:	BOOL;
END_VAR

VAR_INST
	_split	: KOSTAL_AF2024_Core_StringTools.FB_Split_UTF8;
	_resp	: KOSTAL_AF2024_Core_Settings.T_MaxString_UTF8;
	_ETX_1	: STRING(1);
	_ETX_2	: STRING(1);
END_VAR

IF Toggle THEN
	_ETX_1:= Tc2_Standard.LEFT	(_ETX, 1);
	_ETX_2:= Tc2_Standard.RIGHT	(_ETX, 1);
	
	_resp:= KOSTAL_AF2024_Core_StringTools.F_Replace_UTF8(_cmdResponse, _ETX_2, '', -1);
	_split.Split_Delimiter(_resp, _ETX_1);
END_IF

_PrgNumResp:= TO_UINT( _split.Results.line_GET(2));

_catchPrgId:= TRUE;
END_METHOD

METHOD PROTECTED _catchPrgName : BOOL

VAR_INPUT
	Toggle	:	BOOL;
END_VAR

VAR_INST
	_split	: KOSTAL_AF2024_Core_StringTools.FB_Split_UTF8;
	_resp	: KOSTAL_AF2024_Core_Settings.T_MaxString_UTF8;
	_ETX_1	: STRING(1);
	_ETX_2	: STRING(1);
	_str		: KOSTAL_AF2024_Core_Settings.T_MaxString_UTF8;
END_VAR

IF Toggle THEN
	_ETX_1:= Tc2_Standard.LEFT	(_ETX, 1);
	_ETX_2:= Tc2_Standard.RIGHT	(_ETX, 1);
	
	_resp:= KOSTAL_AF2024_Core_StringTools.F_Replace_UTF8(_cmdResponse, _ETX_2, '', -1);
	_split.Split_Delimiter(_resp, _ETX_1);

	_str:= _split.Results.line_GET(2);	//get last entry
END_IF

_split.Split_Delimiter(_str, '/');	//separate optional program location content

_PrgNameResp:= _split.Results.line_GET(_split.Results.NumberOfLines);	//get last entry of string

_catchPrgName:= TRUE;
END_METHOD

METHOD PROTECTED _foundEtx : BOOL
VAR_INPUT
	IN	: KOSTAL_AF2024_Core_Settings.T_MaxString_UTF8;
	OUT	: REFERENCE TO KOSTAL_AF2024_Core_Settings.T_MaxString_UTF8;
END_VAR

VAR
	_OUT	: KOSTAL_AF2024_Core_Settings.T_MaxString_UTF8;
	_pos: INT;
END_VAR

_pos:= Tc2_Standard.FIND(IN, _ETX);

_foundEtx:= _pos <> 0;

IF NOT _foundEtx THEN RETURN;	END_IF

IF NOT __ISVALIDREF(OUT) THEN RETURN;	END_IF

IF _pos = 1 THEN	OUT:= '';
ELSE							OUT:= Tc2_Standard.LEFT(IN, _pos - 1);
END_IF
END_METHOD

METHOD PROTECTED _isCommandAccept : BOOL
VAR_INPUT
	Command	: KOSTAL_AF2024_Core_Settings.T_MaxString;
	Response: KOSTAL_AF2024_Core_Settings.T_MaxString_UTF8;
	Accept	: KOSTAL_AF2024_Core_Settings.T_MaxString_UTF8;
	NoState	: BOOL;
END_VAR

VAR
	_c	: KOSTAL_AF2024_Core_StringTools.FB_Concat;
	_s	: KOSTAL_AF2024_Core_Settings.T_MaxString;
END_VAR

_isCommandAccept:= Tc2_Standard.LEFT(Response, 1) = Accept;//'1';


IF 		_isCommandAccept	THEN	;
ELSE

	_c.Clear();
	_c.addContent(Command);
	_c.addContent(" was not accepted;Errorocode;");
	_c.addContent(TO_WSTRING(Response));
	_s:=  _c.getResult();
	_c.Clear();

	IF NoState	THEN	_State.description:=  _s;	RETURN;	END_IF

	_State.clear();
	_State.description:=  _s;
	_State.fail				:= TRUE;
	_State.finish			:= TRUE;	

END_IF
END_METHOD

METHOD PROTECTED _isPasswordRequest : BOOL
VAR_INPUT
	IN	: KOSTAL_AF2024_Core_Settings.T_MaxString_UTF8;
	NoState	: BOOL;
END_VAR

_isPasswordRequest:= Tc2_Standard.FIND(IN, 'Password:') <> 0;

IF 		_isPasswordRequest	THEN	;
ELSIF NoState							THEN	_State.description:=  "Camera responses no password request";	
ELSE
	_State.clear();
	_State.description:=  "Camera responses no password request";
	_State.fail				:= TRUE;
	_State.finish			:= TRUE;	
END_IF
END_METHOD

METHOD PROTECTED _isUserAccrepted : BOOL
VAR_INPUT
	IN	: KOSTAL_AF2024_Core_Settings.T_MaxString_UTF8;
	NoState	: BOOL;
END_VAR
_isUserAccrepted:= Tc2_Standard.FIND(IN, 'User Logged In') <> 0;

IF 		_isUserAccrepted	THEN	;
ELSIF NoState						THEN	_State.description:= "User login failed";	
ELSE
	_State.clear();
	_State.description:= "User login failed";
	_State.fail				:= TRUE;
	_State.finish			:= TRUE;	
END_IF
END_METHOD

METHOD PROTECTED _isUserRequest : BOOL
VAR_INPUT
	IN	: KOSTAL_AF2024_Core_Settings.T_MaxString_UTF8;
	NoState	: BOOL;
END_VAR
_isUserRequest:= Tc2_Standard.FIND(IN, 'User:') <> 0;

IF 		_isUserRequest	THEN	;
ELSIF NoState					THEN	_State.description:= "Camera responses no User request";	
ELSE
	_State.clear();
	_State.description:= "Camera responses no User request";
	_State.fail				:= TRUE;
	_State.finish			:= TRUE;	
END_IF
END_METHOD

METHOD PROTECTED _isWelcome : BOOL
VAR_INPUT
	IN	: KOSTAL_AF2024_Core_Settings.T_MaxString_UTF8;
	NoState	: BOOL;
END_VAR
_isWelcome:= Tc2_Standard.FIND(IN, 'Welcome') <> 0;

IF 		_isWelcome	THEN	;
ELSIF NoState			THEN	_State.description:= "Camera responses no welcome message";	
ELSE
	_State.clear();
	_State.description:= "Camera responses no welcome message";
	_State.fail				:= TRUE;
	_State.finish			:= TRUE;	
END_IF
END_METHOD

METHOD PROTECTED _SplitData : BOOL
VAR_INST
	_split	:	KOSTAL_AF2024_Core_StringTools.FB_Split_UTF8;
END_VAR

VAR
	_udi: UDINT;
	_dResp: KOSTAL_AF2024_Core_Settings.T_MaxString_UTF8;
	_dResp1: KOSTAL_AF2024_Core_Settings.T_MaxString_UTF8;
	_dResp2: KOSTAL_AF2024_Core_Settings.T_MaxString_UTF8;
END_VAR


//Tc2_Utilities.FindAndDeleteChar(ADR(_dataResponse),	'$R', ADR(_dResp),	SIZEOF(_dResp));
_dResp:= Tc2_Standard.RIGHT(_cmdResponse, Tc2_Standard.LEN(_cmdResponse) - 1);	//remove command part
Tc2_Utilities.FindAndDeleteChar(ADR(_dResp),	'$R', ADR(_dResp1),	SIZEOF(_dResp1));
Tc2_Utilities.FindAndDeleteChar(ADR(_dResp1),	'$N', ADR(_dResp2),	SIZEOF(_dResp2));

_dataResponse:= _dResp2;

_split.Split_Delimiter(_dResp2, ';');

_Data.clear();

FOR _udi:= 1 TO _split.Results.NumberOfLines DO
	_Data.addLine(_split.Results.line_GET(_udi));
END_FOR

_SplitData:= TRUE;
END_METHOD

METHOD PROTECTED _getCommand : KOSTAL_AF2024_Core_Settings.T_MaxString_UTF8

VAR_INPUT
	ID				: E_Command_TcpIp;
	Parameter : KOSTAL_AF2024_Core_Settings.T_MaxString_UTF8;
END_VAR
VAR
	_c	: KOSTAL_AF2024_Core_StringTools.FB_Concat_UTF8;
END_VAR

CASE ID OF

	E_Command_TcpIp.GetInfo		: _getCommand:= 'GI$R$N';			//Returns the system information for the In-Sight vision system.

	E_Command_TcpIp.UserName	: _getCommand:= 'admin$R$N';	//user name.
	E_Command_TcpIp.Password	: _getCommand:= '$R$N';				//password.

	E_Command_TcpIp.SetOnline	: _getCommand:= 'SO1$R$N';		//sets camera to online state.
	E_Command_TcpIp.SetOffline: _getCommand:= 'SO0$R$N';		//sets camera to offline state.

	E_Command_TcpIp.GetOnline	: _getCommand:= 'GO$R$N';			//gets camera online state.
	E_Command_TcpIp.GetPrgId	: _getCommand:= 'GJ$R$N';			//gets camera program (Job) ID.

	E_Command_TcpIp.SetPrgId	: _c.Clear();			//sets camera program (Job) by ID.
															_c.addContent('SJ');
															_c.addContent(Parameter);
															_c.addContent('$R$N');
															_getCommand:= _c.getResult();
															_c.Clear();

	E_Command_TcpIp.SetPrgName	: _c.Clear();			//sets camera program (Job) by Name.
																_c.addContent('LF');
																CASE _PrgLocation OF
																	E_ProgLocation_TcpIp.RamDisk	:	_c.addContent(_STORAGE_RAM_DISK);	_c.addContent('/');
																	E_ProgLocation_TcpIp.SD_Card	:	_c.addContent(_STORAGE_SD_CARD);	_c.addContent('/');
																END_CASE
																_c.addContent(Parameter);
																_c.addContent('$R$N');
																_getCommand:= _c.getResult();
																_c.Clear();
																						
	E_Command_TcpIp.GetPrgName			: _getCommand:= 'GF$R$N';			//gets camera program (Job) name
	E_Command_TcpIp.Trigger					: _getCommand:= 'SW8$R$N';		//triggers camera and wait for result with event 8
	E_Command_TcpIp.GetFormatstring	: _getCommand:= 'GVJob.FormatString$R$N';		//get formatted result(s)
																		
ELSE													_getCommand:= 'UNKNOWN COMMAND';	//return, because no command detected
END_CASE
END_METHOD

METHOD PROTECTED _a3_GetData
VAR
	_split: KOSTAL_AF2024_Core_StringTools.FB_Split_UTF8;
END_VAR

VAR_INST
	_SubStep		: KOSTAL_AF2024_Core_Process.FB_processStep_Flow;
END_VAR

IF _DisableComplexResult THEN	_a3_GetData_DS();
ELSE													_a3_GetData_ETH();
END_IF
END_METHOD

//Get Data over digital signal 
METHOD PROTECTED _a3_GetData_DS
VAR
	_split: KOSTAL_AF2024_Core_StringTools.FB_Split_UTF8;
END_VAR

VAR_INST
	_SubStep		: KOSTAL_AF2024_Core_Process.FB_processStep_Flow;
END_VAR

IF _step.toggle THEN	
	_DigitalSignalRuntimer(IN:= FALSE);	
	_Data.clear();
END_IF

_DigitalSignalRuntimer(IN:= TRUE, PT:= _DigitalSignalRuntime);

IF NOT _DigitalSignalRuntimer.Q THEN

	_State.clear();
	_state.busy	:= TRUE;
	_state.description:= "Wait for digital pass signal";
	
ELSE
	
	IF _DigitalSignal THEN	_Data.addLine('1');
	ELSE										_Data.addLine('0');
	END_IF

	_Step.INC();
	
END_IF
END_METHOD

//Get Data over EtherNet (ETH) 
METHOD PROTECTED _a3_GetData_ETH
VAR
	_split: KOSTAL_AF2024_Core_StringTools.FB_Split_UTF8;
END_VAR

VAR_INST
	_SubStep		: KOSTAL_AF2024_Core_Process.FB_processStep_Flow;
END_VAR

IF _step.toggle THEN
	_Info.clear();

	_state.clear();
	_state.busy:= TRUE;

	_subStep.init();

END_IF


_subStep.Header();


//call command
//===================================================
IF _SubStep.isActive(0)	THEN	_cmd:= _getCommand(E_Command_TcpIp.GetFormatstring, '');
															IF _c1_Send(TRUE, _SubStep.toggle)	THEN	_subStep.INC();	END_IF	
END_IF

//is command accepted?
//===================================================
IF _SubStep.isActive(1)	THEN	IF _c1_Receive(TRUE, _SubStep.toggle)				THEN	_subStep.INC();	END_IF	END_IF
IF _SubStep.isActive(2)	THEN	IF _isCommandAccept("Trigger",_cmdResponse, '1', FALSE)	THEN	_subStep.INC();	END_IF	END_IF

//split data
//===================================================
IF _SubStep.isActive(3)	THEN	IF _SplitData()	THEN	_subStep.INC();	END_IF	END_IF

//finsh
//===================================================
IF _SubStep.isActive(4)	THEN	_Step.INC();	END_IF
END_METHOD

METHOD PROTECTED _a0_stepFail
VAR_INPUT
END_VAR
_connectionInit();
//_isTimeOut(0);

_state.clear();
_state.description:= Tc2_Standard.WCONCAT("Step does not exist: ", INT_TO_WSTRING(_step.actual));
_state.fail		:= TRUE;
_state.finish	:= TRUE;
END_METHOD

METHOD PUBLIC _a0_stepInit
VAR_INPUT
END_VAR

//Overwrite base method

IF _Init OR_ELSE (_THIS_CALLED <> _THIS_IN_PROCESS AND _step.actual > 0) THEN 

	_step.init();
	_Init:= FALSE;	

	_ConnectionInit();
	
END_IF
END_METHOD

METHOD PROTECTED _a1_failure
VAR_INPUT
	lState	: KOSTAL_AF2024_Core_Process.I_T_plcState;
	Toggle	: BOOL;
END_VAR

VAR
	_obj	: KOSTAL_AF2024_Core_Process.I_T_plcState;
END_VAR

VAR_INST
	_lState	: KOSTAL_AF2024_Core_Process.T_plcState;
END_VAR

IF lState <> 0 AND_THEN __QUERYINTERFACE(lState, _obj) AND_THEN _obj <> 0 THEN
	
	IF Toggle THEN _lState.CopyFrom(lState);	END_IF

	_State.CopyFrom(_lState);

END_IF
END_METHOD

METHOD PROTECTED _a1_Finish

IF _step.toggle THEN

	_connectionInit();

END_IF

_State.clear();
_State.finish	:= TRUE;
_State.pass		:= TRUE;
END_METHOD

METHOD PROTECTED _a1_Idle

_state.clear();

_THIS_IN_PROCESS:= _E_THIS_TcpIp.Idle;

_ConnectionInit();

IF 	_cmdSocket.bBusy THEN

	_state.busy:= TRUE;
	_state.description:= "command socket is busy, please wait...";
	
ELSIF _cmdSend.bBusy THEN

	_state.busy:= TRUE;
	_state.description:= "command send is busy, please wait...";

	
ELSIF _cmdReceive.bBusy THEN

	_state.busy:= TRUE;
	_state.description:= "command receive is busy, please wait...";


ELSIF _THIS_CALLED = _E_THIS_TcpIp.Idle THEN

	_state.ready:= TRUE;

ELSIF _THIS_CALLED = _E_THIS_TcpIp.GetInfo THEN

	_THIS_IN_PROCESS:= _THIS_CALLED;

	_state.busy:= TRUE;

	_cmdReceivedString:= '';
	_cmdReceivedPartly:= '';

	_Info.Clear();
	
	_step.set(_ADDRESS_GetInfo);
	
	
ELSIF _THIS_CALLED = _E_THIS_TcpIp.Trigger THEN

	_THIS_IN_PROCESS:= _THIS_CALLED;

	_state.busy:= TRUE;

	_cmdReceivedString:= '';
	_cmdReceivedPartly:= '';


	_Data.clear();
	
	_step.set(_ADDRESS_Trigger);

	
ELSIF _THIS_CALLED = _E_THIS_TcpIp.TriggerPrgNo THEN

	_THIS_IN_PROCESS:= _THIS_CALLED;

	_state.busy:= TRUE;

	_cmdReceivedString:= '';
	_cmdReceivedPartly:= '';

	_Data.clear();

	_step.set(_ADDRESS_TriggerPrgNum);

	
ELSIF _THIS_CALLED = _E_THIS_TcpIp.TriggerPrgName THEN

	_THIS_IN_PROCESS:= _THIS_CALLED;

	_state.busy:= TRUE;

	_cmdReceivedString:= '';
	_cmdReceivedPartly:= '';

	_Data.clear();

	_step.set(_ADDRESS_TriggerPrgName);

ELSIF _THIS_CALLED = _E_THIS_TcpIp.SetProgramId THEN

	_THIS_IN_PROCESS:= _THIS_CALLED;

	_state.busy:= TRUE;

	_cmdReceivedString:= '';
	_cmdReceivedPartly:= '';

	_step.set(_ADDRESS_SetPrgNum);
	

ELSIF _THIS_CALLED = _E_THIS_TcpIp.SetProgramName THEN

	_THIS_IN_PROCESS:= _THIS_CALLED;

	_state.busy:= TRUE;

	_cmdReceivedString:= '';
	_cmdReceivedPartly:= '';

	_step.set(_ADDRESS_SetPrgName);
	

ELSIF _THIS_CALLED = _E_THIS_TcpIp.GetProgramId THEN

	_THIS_IN_PROCESS:= _THIS_CALLED;

	_state.busy:= TRUE;

	_cmdReceivedString:= '';
	_cmdReceivedPartly:= '';

	_step.set(_ADDRESS_GetPrgNum);
	

ELSIF _THIS_CALLED = _E_THIS_TcpIp.GetProgramName THEN

	_THIS_IN_PROCESS:= _THIS_CALLED;

	_state.busy:= TRUE;

	_cmdReceivedString:= '';
	_cmdReceivedPartly:= '';

	_step.set(_ADDRESS_GetPrgName);
	
	
ELSIF _THIS_CALLED = _E_THIS_TcpIp.Idle THEN

	_state.clear();
	_state.ready:= TRUE;
		
ELSE

	_State.clear();
	_State.finish:= TRUE;
	_State.fail:= TRUE;
	_State.description:= "Unknown command detected";

END_IF
END_METHOD

METHOD PROTECTED _a2_Login

VAR_INST
	_SubStep		: KOSTAL_AF2024_Core_Process.FB_processStep_Flow;
	_hasUserRequest	: BOOL;
END_VAR

IF _step.toggle THEN

	_state.clear();
	_state.busy:= TRUE;

	_subStep.init();
	
END_IF


_subStep.Header();

//Initialize/disconnect sockets	
//===================================================
IF _SubStep.isActive(0)	THEN	IF _c1_Socket(FALSE) THEN	_subStep.INC();	END_IF	END_IF
IF _SubStep.isActive(1)	THEN	IF _c1_Socket(TRUE) THEN	_subStep.INC();	END_IF	END_IF


//connect and is welcome? and save has user request?
//===================================================
IF _SubStep.isActive(2)	THEN	IF _c1_Receive(TRUE, _SubStep.toggle)	THEN _SubStep.INC();	END_IF	END_IF

IF _SubStep.isActive(3)	THEN	
	IF _SubStep.toggle THEN _hasUserRequest:= _isUserRequest(_cmdResponse, TRUE);	END_IF
	IF _isWelcome(_cmdResponse, FALSE)	THEN _SubStep.INC();	END_IF
END_IF
	
//get user request if not exist in first call
//===================================================
IF _SubStep.isActive(4)	THEN	
	IF NOT _hasUserRequest THEN
		IF _c1_Receive(TRUE, _SubStep.toggle)	THEN _SubStep.INC();	END_IF
	ELSE	_SubStep.INC();
	END_IF
END_IF
	
//is user request
//===================================================
IF _SubStep.isActive(5)	THEN	
	IF NOT _hasUserRequest THEN	IF _isUserRequest(_cmdResponse, FALSE)	THEN	_subStep.INC();	END_IF
	ELSE 												_SubStep.INC();
	END_IF
END_IF

//send user name
//===================================================
IF _SubStep.isActive(6)	THEN	_cmd:= _getCommand(E_Command_TcpIp.UserName, '');
															IF _c1_Send(TRUE, _SubStep.toggle)	THEN	_subStep.INC();	END_IF	
END_IF


//is password requested?
//===================================================
IF _SubStep.isActive(7)	THEN	IF _c1_Receive(TRUE, _SubStep.toggle)	THEN	_subStep.INC();	END_IF	END_IF
IF _SubStep.isActive(8)	THEN	_c1_Socket(TRUE);	IF _isPasswordRequest(_cmdResponse, FALSE)				THEN	_subStep.INC();	END_IF	END_IF
	
//send password
//===================================================
IF _SubStep.isActive(9)	THEN	_cmd:= _getCommand(E_Command_TcpIp.Password, '');
															IF _c1_Send(TRUE, _SubStep.toggle)	THEN	_subStep.INC();	END_IF	
END_IF

//is login accepted?
//===================================================
IF _SubStep.isActive(10)	THEN	IF _c1_Receive(TRUE, _SubStep.toggle)	THEN	_subStep.INC();	END_IF	END_IF
IF _SubStep.isActive(11)	THEN	_c1_Socket(TRUE);	IF _isUserAccrepted(_cmdResponse, FALSE)			THEN	_subStep.INC();	END_IF	END_IF

//connection successful
//===================================================
IF _SubStep.isActive(12)	THEN	_c1_Socket(TRUE);	 _Step.INC();	END_IF
END_METHOD

METHOD PROTECTED _a3_GetInfo
VAR
	_splitLine: KOSTAL_AF2024_Core_StringTools.FB_Split_UTF8;
	_split		: KOSTAL_AF2024_Core_StringTools.FB_Split_UTF8;
	_udi			: UDINT;
END_VAR

VAR_INST
	_SubStep	: KOSTAL_AF2024_Core_Process.FB_processStep_Flow;
	_InformationNotConclusive	: BOOL;
	_resp			: KOSTAL_AF2024_Core_Settings.T_MaxString_UTF8;
	_resp1		: KOSTAL_AF2024_Core_Settings.T_MaxString_UTF8;
END_VAR

IF _step.toggle THEN
	_Info.clear();

	_state.clear();
	_state.busy:= TRUE;

	_subStep.init();


END_IF


_subStep.Header();


//call command
//===================================================
IF _SubStep.isActive(0)	THEN	_cmd:= _getCommand(E_Command_TcpIp.GetInfo, '');
															IF _c1_Send(TRUE, _SubStep.toggle)	THEN	_subStep.INC();	END_IF	
END_IF

//is command accepted?
//===================================================
IF _SubStep.isActive(1)	THEN	IF _c1_Receive(TRUE, _SubStep.toggle)				THEN	_subStep.INC();	END_IF	END_IF
//IF _SubStep.isActive(2)	THEN	_c1_Socket(TRUE); IF _isCommandAccept("GetInfo",_cmdResponse)	THEN	_subStep.INC();	_Line:= 0;	END_IF	END_IF

//get line
//===================================================
//IF _SubStep.isActive(3)	THEN	(*_AddressLoopHeader:= _SubStep.actual;*)
//															IF _c1_Receive(TRUE, _SubStep.toggle) THEN	_subStep.INC();	(*_Line:= _Line + 1;*)	END_IF	
//END_IF


//parse line
//===================================================
IF _SubStep.isActive(2)	THEN	
	
		
	IF _SubStep.toggle THEN	_c1_Socket(FALSE);	_splitLine.Split_Delimiter(_cmdResponse, '$0D');	END_IF	

	IF NOT _isCommandAccept("GetInfo", _splitLine.Results.line_GET(1), '1', FALSE)	THEN	;

	ELSE
	
		_InformationNotConclusive:= FALSE;
		
		FOR _udi:= 2 TO _splitLine.Results.NumberOfLines - 1 DO

			_split.Clear();	
			_split.Split_Delimiter(_splitLine.Results.line_GET(_udi), ':');	
			_resp1:= Tc2_Utilities.F_LTrim(_split.Results.line_GET(2)); 
			Tc2_Utilities.FindAndDeleteChar(ADR(_resp1), '$0A', ADR(_resp), SIZEOF(_resp));	
			
			IF 		Tc2_Standard.FIND (_split.Results.line_GET(1), 'Serial') <> 0 			THEN	_Info.SerialNumber			:= _resp;
			ELSIF Tc2_Standard.FIND (_split.Results.line_GET(1), 'Application') <> 0	THEN	_Info.ApplicationVersion:= _resp;
			ELSIF Tc2_Standard.FIND (_split.Results.line_GET(1), 'Monitor') <> 0			THEN	_Info.MonitorVersion		:= _resp;
			ELSIF Tc2_Standard.FIND (_split.Results.line_GET(1), 'MAC') <> 0					THEN	_Info.MonitorVersion 		:= _catchMacId(_resp);
			ELSIF Tc2_Standard.FIND (_split.Results.line_GET(1), 'Date') <> 0					THEN	_Info.DateOfBuild				:= _resp;
			ELSE	_InformationNotConclusive:= TRUE;	
			END_IF
			
		END_FOR
		
		_SubStep.INC();
		
	END_IF
END_IF

//finish
//===================================================
IF _SubStep.isActive(3)	THEN

	IF _InformationNotConclusive THEN
				_State.clear();
				_State.description:= "Information is not conclusive";
				_State.fail	:= TRUE;
				_State.finish:= TRUE;	

	ELSE	_Step.INC();
	END_IF
		
END_IF
END_METHOD

METHOD PROTECTED _a3_GetPrgId

VAR_INST
	_SubStep		: KOSTAL_AF2024_Core_Process.FB_processStep_Flow;
	_AddressFinish 	: INT:= 10;
END_VAR

IF _step.toggle THEN
	_PrgNumResp:= 16#FFFF;
	
	_state.clear();
	_state.busy:= TRUE;

	_subStep.init();

END_IF


_subStep.Header();

//call command
//===================================================
IF _SubStep.isActive(0)	THEN	_cmd:= _getCommand(E_Command_TcpIp.GetPrgId, '');
															IF _c1_Send(TRUE, _SubStep.toggle)	THEN	_subStep.INC();	END_IF	
END_IF

//is command accepted?
//===================================================
IF _SubStep.isActive(1)	THEN	IF _c1_Receive(TRUE, _SubStep.toggle)				THEN	_subStep.INC();	END_IF	END_IF
IF _SubStep.isActive(2)	THEN	IF _isCommandAccept("GetPrgId",_cmdResponse, '1', TRUE)	THEN		_subStep.INC(); ELSE 	_subStep.set(_AddressFinish); END_IF	END_IF
IF _SubStep.isActive(3)	THEN	IF _catchPrgId(_SubStep.toggle)													THEN	_subStep.set(_AddressFinish);	END_IF	END_IF


//finsh
//===================================================
IF _SubStep.isActive(_AddressFinish)	THEN	_Step.INC();	END_IF
END_METHOD

METHOD PROTECTED _a3_GetPrgName

VAR_INST
	_SubStep				: KOSTAL_AF2024_Core_Process.FB_processStep_Flow;
	_AddressFinish 	: INT:= 10;
END_VAR

IF _step.toggle THEN
	_PrgNameResp:= '';
	
	_state.clear();
	_state.busy:= TRUE;

	_subStep.init();

END_IF


_subStep.Header();

//call command
//===================================================
IF _SubStep.isActive(0)	THEN	_cmd:= _getCommand(E_Command_TcpIp.GetPrgName, '');
															IF _c1_Send(TRUE, _SubStep.toggle)	THEN	_subStep.INC();	END_IF	
END_IF

//is command accepted?
//===================================================
IF _SubStep.isActive(1)	THEN	IF _c1_Receive(TRUE, _SubStep.toggle)					THEN	_subStep.INC();	END_IF	END_IF
IF _SubStep.isActive(2)	THEN	IF _isCommandAccept("GetPrgName",_cmdResponse, '1', TRUE)	THEN	_subStep.INC();	ELSE	_subStep.set(_AddressFinish);	END_IF	END_IF
IF _SubStep.isActive(3)	THEN	IF _catchPrgName(_SubStep.toggle)													THEN	_subStep.set(_AddressFinish);	END_IF	END_IF


//finsh
//===================================================
IF _SubStep.isActive(_AddressFinish)	THEN	_Step.INC();	END_IF
END_METHOD

METHOD PROTECTED _a3_SetOffline

VAR_INPUT
	Enable	: BOOL;
END_VAR


VAR_INST
	_SubStep		: KOSTAL_AF2024_Core_Process.FB_processStep_Flow;
END_VAR
IF _step.toggle THEN

	_state.clear();
	_state.busy:= TRUE;

	_subStep.init();

END_IF

_subStep.Header();

//analyse enable bit
//===================================================
IF _SubStep.isActive(0)	THEN	IF NOT Enable THEN	_Step.INC();	ELSE	_SubStep.INC();	END_IF	END_IF

//call command
//===================================================
IF _SubStep.isActive(1)	THEN	_cmd:= _getCommand(E_Command_TcpIp.SetOffline, '');
	IF _c1_Send(TRUE, _SubStep.toggle)	THEN	_subStep.INC();	END_IF	
END_IF

//is command accepted?
//===================================================
IF _SubStep.isActive(2)	THEN	IF _c1_Receive(TRUE, _SubStep.toggle)							THEN	_subStep.INC();	END_IF	END_IF
IF _SubStep.isActive(3)	THEN	IF _isCommandAccept("SetOffline",_cmdResponse, '1', FALSE)	THEN	_subStep.INC();	END_IF	END_IF

//finsh
//===================================================
IF _SubStep.isActive(4)	THEN	_Step.INC();	END_IF
END_METHOD

METHOD PROTECTED _a3_SetOnline

VAR_INST
	_SubStep		: KOSTAL_AF2024_Core_Process.FB_processStep_Flow;
END_VAR

IF _step.toggle THEN

	_state.clear();
	_state.busy:= TRUE;

	_subStep.init();

END_IF

_subStep.Header();

//call command
//===================================================
IF _SubStep.isActive(0)	THEN	_cmd:= _getCommand(E_Command_TcpIp.SetOnline, '');
	IF _c1_Send(TRUE, _SubStep.toggle)	THEN	_subStep.INC();	END_IF	
END_IF

//is command accepted?
//===================================================
IF _SubStep.isActive(1)	THEN	IF _c1_Receive(TRUE, _SubStep.toggle)							THEN	_subStep.INC();	END_IF	END_IF
IF _SubStep.isActive(2)	THEN	IF _isCommandAccept("SetOnline",_cmdResponse, '1', FALSE)	THEN	_subStep.INC();	END_IF	END_IF

//finsh
//===================================================
IF _SubStep.isActive(3)	THEN	_Step.INC();	END_IF
END_METHOD

METHOD PROTECTED _a3_SetReqPrgById

VAR_INPUT
	Enable	: BOOL;
END_VAR


VAR_INST
	_SubStep		: KOSTAL_AF2024_Core_Process.FB_processStep_Flow;
END_VAR
IF _step.toggle THEN

	_state.clear();
	_state.busy:= TRUE;

	_subStep.init();

END_IF

_subStep.Header();

//analyse the enable bit
//===================================================
IF _SubStep.isActive(0)	THEN	IF NOT Enable THEN	_Step.INC();	ELSE	_SubStep.INC();	END_IF	END_IF

//call command
//===================================================
IF _SubStep.isActive(1)	THEN	_cmd:= _getCommand(E_Command_TcpIp.SetPrgId, TO_STRING(_PrgNum));
	IF _c1_Send(TRUE, _SubStep.toggle)	THEN	_subStep.INC();	END_IF	
END_IF

//is command accepted?
//===================================================
IF _SubStep.isActive(2)	THEN	IF _c1_Receive(TRUE, _SubStep.toggle)									THEN	_subStep.INC();	END_IF	END_IF
IF _SubStep.isActive(3)	THEN	IF _isCommandAccept("SetreqPrg",_cmdResponse, '1', FALSE)	THEN _PrgNumResp:= _PrgNum;	_subStep.INC();	END_IF	END_IF

//finsh
//===================================================
IF _SubStep.isActive(4)	THEN	_Step.INC();	END_IF
END_METHOD

METHOD PROTECTED _a3_SetReqPrgByName

VAR_INPUT
	Enable	: BOOL;
END_VAR


VAR_INST
	_SubStep		: KOSTAL_AF2024_Core_Process.FB_processStep_Flow;
END_VAR
IF _step.toggle THEN

	_state.clear();
	_state.busy:= TRUE;

	_subStep.init();

END_IF

_subStep.Header();

//analyse the enable bit
//===================================================
IF _SubStep.isActive(0)	THEN	IF NOT Enable THEN	_Step.INC();	ELSE	_SubStep.INC();	END_IF	END_IF

//call command
//===================================================
IF _SubStep.isActive(1)	THEN	_cmd:= _getCommand(E_Command_TcpIp.SetPrgName, _PrgName);
	IF _c1_Send(TRUE, _SubStep.toggle)	THEN	_subStep.INC();	END_IF	
END_IF

//is command accepted?
//===================================================
IF _SubStep.isActive(2)	THEN	IF _c1_Receive(TRUE, _SubStep.toggle)									THEN	_subStep.INC();	END_IF	END_IF
IF _SubStep.isActive(3)	THEN	IF _isCommandAccept("SetreqPrg",_cmdResponse, '1', FALSE)	THEN	_PrgNameResp:= _PrgName;	_subStep.INC();	END_IF	END_IF

//finsh
//===================================================
IF _SubStep.isActive(4)	THEN	_Step.INC();	END_IF
END_METHOD

METHOD PROTECTED _a3_Trigger
VAR
	_split: KOSTAL_AF2024_Core_StringTools.FB_Split_UTF8;
END_VAR

VAR_INST
	_SubStep		: KOSTAL_AF2024_Core_Process.FB_processStep_Flow;
END_VAR

IF _step.toggle THEN
	_Info.clear();

	_state.clear();
	_state.busy:= TRUE;

	_subStep.init();

END_IF


_subStep.Header();

//call command
//===================================================
IF _SubStep.isActive(0)	THEN	_cmd:= _getCommand(E_Command_TcpIp.Trigger, '');
															IF _c1_Send(TRUE, _SubStep.toggle)	THEN	_subStep.INC();	END_IF	
END_IF

//is command accepted?
//===================================================
IF _SubStep.isActive(1)	THEN	IF _c1_Receive(TRUE, _SubStep.toggle)								THEN	_subStep.INC();	END_IF	END_IF
IF _SubStep.isActive(2)	THEN	IF _isCommandAccept("Trigger",_cmdResponse, '1', FALSE)	THEN	_subStep.INC();	END_IF	END_IF

//finsh
//===================================================
IF _SubStep.isActive(3)	THEN	_Step.INC();	END_IF
END_METHOD

(*
Decription
==========
*)
METHOD PROTECTED _FBmain

//_d1_Server();

_a0_stepInit();

_step.Header();

IF _Step.isActive(0)	THEN	_a1_Idle();	END_IF
	
//Get Info
IF _Step.isActive(_ADDRESS_GetInfo)			THEN	_a2_Login();		END_IF
IF _Step.isActive(_ADDRESS_GetInfo + 1)	THEN	_a3_GetInfo();	END_IF
IF _Step.isActive(_ADDRESS_GetInfo + 2)	THEN	_a1_Finish();		END_IF

//trigger only
IF _Step.isActive(_ADDRESS_Trigger)			THEN	_a2_Login();			END_IF
IF _Step.isActive(_ADDRESS_Trigger + 1)	THEN	_a3_Trigger();		END_IF
IF _Step.isActive(_ADDRESS_Trigger + 2)	THEN	_a3_GetData();		END_IF
IF _Step.isActive(_ADDRESS_Trigger + 3)	THEN	_a1_Finish();			END_IF


//trigger prg num (Job ID)
IF _Step.isActive(_ADDRESS_TriggerPrgNum)			THEN	_a2_Login();			END_IF
IF _Step.isActive(_ADDRESS_TriggerPrgNum + 1)	THEN	_a3_GetPrgId();		END_IF
IF _Step.isActive(_ADDRESS_TriggerPrgNum + 2)	THEN	_a3_SetOffline(_PrgNum <> _PrgNumResp);			END_IF
IF _Step.isActive(_ADDRESS_TriggerPrgNum + 3)	THEN	_a3_SetReqPrgById(_PrgNum <> _PrgNumResp);	END_IF
IF _Step.isActive(_ADDRESS_TriggerPrgNum + 4)	THEN	_a3_SetOnline();	END_IF
IF _Step.isActive(_ADDRESS_TriggerPrgNum + 5)	THEN	_a3_Trigger();		END_IF
IF _Step.isActive(_ADDRESS_TriggerPrgNum + 6)	THEN	_a3_GetData();		END_IF
IF _Step.isActive(_ADDRESS_TriggerPrgNum + 7)	THEN	_a1_Finish();			END_IF

//trigger prg name (Job File Name)
IF _Step.isActive(_ADDRESS_TriggerPrgName)			THEN	_a2_Login();			END_IF
IF _Step.isActive(_ADDRESS_TriggerPrgName + 1)	THEN	_a3_GetPrgName();	END_IF
IF _Step.isActive(_ADDRESS_TriggerPrgName + 2)	THEN	_a3_SetOffline(_PrgName <> _PrgNameResp);				END_IF
IF _Step.isActive(_ADDRESS_TriggerPrgName + 3)	THEN	_a3_SetReqPrgByName(_PrgName <> _PrgNameResp);	END_IF
IF _Step.isActive(_ADDRESS_TriggerPrgName + 4)	THEN	_a3_SetOnline();	END_IF
IF _Step.isActive(_ADDRESS_TriggerPrgName + 5)	THEN	_a3_Trigger();		END_IF
IF _Step.isActive(_ADDRESS_TriggerPrgName + 6)	THEN	_a3_GetData();		END_IF
IF _Step.isActive(_ADDRESS_TriggerPrgName + 7)	THEN	_a1_Finish();			END_IF

//set prg num (Job ID)
IF _Step.isActive(_ADDRESS_SetPrgNum)			THEN	_a2_Login();							END_IF
IF _Step.isActive(_ADDRESS_SetPrgNum + 1)	THEN	_a3_SetOffline(TRUE);			END_IF
IF _Step.isActive(_ADDRESS_SetPrgNum + 2)	THEN	_a3_SetReqPrgById(TRUE);	END_IF
IF _Step.isActive(_ADDRESS_SetPrgNum + 3)	THEN	_a3_SetOnline();					END_IF
IF _Step.isActive(_ADDRESS_SetPrgNum + 4)	THEN	_a1_Finish();							END_IF

//set prg name (Job file name)
IF _Step.isActive(_ADDRESS_SetPrgName)			THEN	_a2_Login();								END_IF
IF _Step.isActive(_ADDRESS_SetPrgName + 1)	THEN	_a3_SetOffline(TRUE);				END_IF
IF _Step.isActive(_ADDRESS_SetPrgName + 2)	THEN	_a3_SetReqPrgByName(TRUE);	END_IF
IF _Step.isActive(_ADDRESS_SetPrgName + 3)	THEN	_a3_SetOnline();						END_IF
IF _Step.isActive(_ADDRESS_SetPrgName + 4)	THEN	_a1_Finish();								END_IF


//get Program ID
IF _Step.isActive(_ADDRESS_GetPrgNum)			THEN	_a2_Login();		END_IF
IF _Step.isActive(_ADDRESS_GetPrgNum + 1)	THEN	_a3_GetPrgId();	END_IF
IF _Step.isActive(_ADDRESS_GetPrgNum + 2)	THEN	_a1_Finish();		END_IF

//get Program Name
IF _Step.isActive(_ADDRESS_GetPrgName)			THEN	_a2_Login();			END_IF
IF _Step.isActive(_ADDRESS_GetPrgName + 1)	THEN	_a3_GetPrgName();	END_IF
IF _Step.isActive(_ADDRESS_GetPrgName + 2)	THEN	_a1_Finish();			END_IF


IF _Step.NotFound()	THEN _a0_stepFail();	END_IF
END_METHOD

METHOD Ex_GetInfo : BOOL
VAR_INPUT
	Info	: I_T_Info_TcpIp;
END_VAR

VAR
	_obj	: I_T_Info_TcpIp;
END_VAR
;

IF _THIS_CALLED = _E_THIS_TcpIp.Idle THEN

	_THIS_CALLED:= _E_THIS_TcpIp.GetInfo;

	_FBmain();

	Ex_GetInfo:= _THIS_CALLED = _THIS_IN_PROCESS;

	IF Ex_GetInfo AND_THEN __QUERYINTERFACE(Info, _obj) AND_THEN _obj <> 0 THEN Info:= _Info;	END_IF
 
ELSE

	Ex_GetInfo:= FALSE;
	
END_IF
END_METHOD

METHOD Ex_GetProgamNumber : BOOL
VAR_INPUT
	Number	: REFERENCE TO UINT;
END_VAR
IF _THIS_CALLED = _E_THIS_TcpIp.Idle THEN

	_THIS_CALLED:= _E_THIS_TcpIp.GetProgramId;

	_FBmain();

	Ex_GetProgamNumber:= _THIS_CALLED = _THIS_IN_PROCESS;
	
	IF Ex_GetProgamNumber AND_THEN __ISVALIDREF(Number) THEN Number:= _PrgNumResp;	END_IF

ELSE
	
	Ex_GetProgamNumber:= FALSE;
 
END_IF
END_METHOD

METHOD Ex_GetProgramName : BOOL
VAR_INPUT
	Name	: REFERENCE TO KOSTAL_AF2024_Core_Settings.T_MaxString_UTF8;
END_VAR
IF _THIS_CALLED = _E_THIS_TcpIp.Idle THEN

	_THIS_CALLED:= _E_THIS_TcpIp.GetProgramName;

	_FBmain();

	Ex_GetProgramName:= _THIS_CALLED = _THIS_IN_PROCESS;
	
	IF Ex_GetProgramName AND_THEN __ISVALIDREF(Name) THEN Name:= _PrgNameResp;	END_IF
	
ELSE
	
	Ex_GetProgramName:= FALSE;
 
END_IF
END_METHOD

METHOD Ex_SetProgramName : BOOL
VAR_INPUT
	Name	: KOSTAL_AF2024_Core_Settings.T_MaxString_UTF8;
END_VAR
IF _THIS_CALLED = _E_THIS_TcpIp.Idle THEN

	_THIS_CALLED:= _E_THIS_TcpIp.SetProgramName;

	_PrgName:= Name;

	_FBmain();

	Ex_SetProgramName:= _THIS_CALLED = _THIS_IN_PROCESS;
	
ELSE
	
	Ex_SetProgramName:= FALSE;
 
END_IF
END_METHOD

METHOD Ex_SetProgramNumber : BOOL
VAR_INPUT
	ProgramNumber	: UINT;
END_VAR
IF _THIS_CALLED = _E_THIS_TcpIp.Idle THEN

	_THIS_CALLED:= _E_THIS_TcpIp.SetProgramId;

	_PrgNum:= ProgramNumber;

	_FBmain();

	Ex_SetProgramNumber:= _THIS_CALLED = _THIS_IN_PROCESS;
	
ELSE
	
	Ex_SetProgramNumber:= FALSE;
 
END_IF
END_METHOD

METHOD Ex_Trigger : BOOL
;

IF _THIS_CALLED = _E_THIS_TcpIp.Idle THEN

	_THIS_CALLED:= _E_THIS_TcpIp.Trigger;

	_FBmain();

	Ex_Trigger:= _THIS_CALLED = _THIS_IN_PROCESS;

ELSE

	Ex_Trigger:= FALSE;
	
END_IF
END_METHOD

METHOD Ex_Trigger_ProgName : BOOL
VAR_INPUT
	ProgName	: KOSTAL_AF2024_Core_Settings.T_MaxString_UTF8;
END_VAR

IF _THIS_CALLED = _E_THIS_TcpIp.Idle THEN

	_THIS_CALLED:= _E_THIS_TcpIp.TriggerPrgName;
	
	_PrgName:= ProgName;
	
	_FBmain();

	Ex_Trigger_ProgName:= _THIS_CALLED = _THIS_IN_PROCESS;

ELSE

	Ex_Trigger_ProgName:= FALSE;
	
END_IF
END_METHOD

METHOD Ex_Trigger_ProgramNumber : BOOL
VAR_INPUT
	ProgramNumber	: UINT;
END_VAR
IF _THIS_CALLED = _E_THIS_TcpIp.Idle THEN

	_THIS_CALLED:= _E_THIS_TcpIp.TriggerPrgNo;
	
	_PrgNum:= ProgramNumber;
	
	_FBmain();

	Ex_Trigger_ProgramNumber:= _THIS_CALLED = _THIS_IN_PROCESS;

ELSE

	Ex_Trigger_ProgramNumber:= FALSE;
	
END_IF
END_METHOD

(*
Description
===========
| TCP/IP port of the barcode reader
*)
PROPERTY PUBLIC CommandPort : UDINT
GET


CommandPort:= _CmdPort;
END_GET
SET

IF CommandPort = UDINT#0 THEN	_CmdPort:= _CMD_PORT_DEFAULT;
ELSE													_CmdPort:= CommandPort;
END_IF
END_SET
END_PROPERTY

PROPERTY PUBLIC CommandTimeOut : TIME
GET

CommandTimeOut:= _cmdTimeOut;
END_GET
SET

IF CommandTimeOut > T#5S THEN	_cmdTimeOut:= CommandTimeOut;	ELSE _cmdTimeOut:= _DEFAULT_TIMEOUT;	END_IF
END_SET
END_PROPERTY

(*
Description
===========
| IP address of the barcode reader
*)
PROPERTY PUBLIC IP : STRING
GET


IP:= _IP;
END_GET
SET

_IP:= IP;
END_SET
END_PROPERTY

PROPERTY PUBLIC Data : KOSTAL_AF2024_Core_ListOf.I_ListOfString_UTF8
GET

Data:= _Data;
END_GET
END_PROPERTY

//Waiting time before the digital signal is analyzed.
PROPERTY PUBLIC DigitalSignalRuntime : TIME
GET

DigitalSignalRuntime:= _DigitalSignalRuntime;
END_GET
SET

_DigitalSignalRuntime:= DigitalSignalRuntime;
END_SET
END_PROPERTY

PROPERTY PUBLIC DisableComplexResult : BOOL
GET

DisableComplexResult:= _DisableComplexResult;
END_GET
SET

_DisableComplexResult:= DisableComplexResult;
END_SET
END_PROPERTY

PROPERTY PUBLIC Info : I_T_Info_TcpIp
GET

Info:= _Info;
END_GET
END_PROPERTY

PROPERTY PUBLIC ProgLocation : E_ProgLocation_TcpIp
GET

ProgLocation:= _PrgLocationResp;
END_GET
SET

_PrgLocation:= ProgLocation;
END_SET
END_PROPERTY

PROPERTY ResultPass : BOOL
GET

ResultPass:= _Data.line_GET(1) = '1';	//Tc2_Standard.LEFT(_cmdResponse,1) = '1';
END_GET
END_PROPERTY

PROPERTY State : KOSTAL_AF2024_Drivers_Camera_I_Camera.KOSTAL_AF2024_Core_Process.I_T_plcState
GET

State:= _State;
END_GET
END_PROPERTY

(*
Decription
==========
| To be called cyclicly, e.g. in DeviceDefine
*)
METHOD PUBLIC FBmain
VAR_INPUT
END_VAR

IF _THIS_CALLED = _E_THIS_TcpIp.Idle THEN
	_FBmain();
END_IF

_THIS_CALLED:= _E_THIS_TcpIp.Idle;
END_METHOD

END_FUNCTION_BLOCK

// TcpIp/I_InSight_TcpIp
INTERFACE I_InSight_TcpIp EXTENDS KOSTAL_AF2024_Drivers_Camera_I_Camera.I_Camera

METHOD Ex_GetInfo : BOOL
VAR_INPUT
	Info	: I_T_Info_TcpIp;
END_VAR
END_METHOD

METHOD Ex_GetProgamNumber : BOOL
VAR_INPUT
	Number	: REFERENCE TO UINT;
END_VAR
END_METHOD

METHOD Ex_GetProgramName : BOOL
VAR_INPUT
	Name	: REFERENCE TO KOSTAL_AF2024_Core_Settings.T_MaxString_UTF8;
END_VAR
END_METHOD

METHOD Ex_SetProgramName : BOOL
VAR_INPUT
	Name	: KOSTAL_AF2024_Core_Settings.T_MaxString_UTF8;
END_VAR
END_METHOD

METHOD Ex_Trigger_ProgName : BOOL
VAR_INPUT
	ProgName	: KOSTAL_AF2024_Core_Settings.T_MaxString_UTF8;
END_VAR
END_METHOD

(*
Description
===========
| TCP/IP port of the barcode reader
*)
PROPERTY PUBLIC CommandPort : UDINT
GET
END_GET
SET
END_SET
END_PROPERTY

PROPERTY PUBLIC CommandTimeOut : TIME
GET
END_GET
SET
END_SET
END_PROPERTY

(*
Description
===========
| IP address of the barcode reader
*)
PROPERTY PUBLIC IP : STRING
GET
END_GET
SET
END_SET
END_PROPERTY

PROPERTY PUBLIC Data : KOSTAL_AF2024_Core_ListOf.I_ListOfString_UTF8
GET
END_GET
END_PROPERTY

//Waiting time before the digital signal is analyzed.
PROPERTY PUBLIC DigitalSignalRuntime : TIME
GET
END_GET
SET
END_SET
END_PROPERTY

PROPERTY PUBLIC DisableComplexResult : BOOL
GET
END_GET
SET
END_SET
END_PROPERTY

PROPERTY PUBLIC Info : I_T_Info_TcpIp
GET
END_GET
END_PROPERTY

PROPERTY PUBLIC ProgLocation : E_ProgLocation_TcpIp
GET
END_GET
SET
END_SET
END_PROPERTY

END_INTERFACE

// TcpIp/FB_InSight_VisionSuite_TcpIp
FUNCTION_BLOCK PUBLIC FB_InSight_VisionSuite_TcpIp EXTENDS FB_InSight_Explorer_TcpIp
VAR
	_sheetName	: KOSTAL_AF2024_Core_Settings.T_MaxString_UTF8 := 'AF_2024';
END_VAR

//cameras with InSigtVisionSuite sends MAC ID with ':'
METHOD PROTECTED _catchMacId : KOSTAL_AF2024_Core_Settings.T_MaxString_UTF8
VAR_INPUT
	IN	: KOSTAL_AF2024_Core_Settings.T_MaxString_UTF8;
END_VAR

VAR
	_IN		: KOSTAL_AF2024_Core_Settings.T_MaxString_UTF8;
	_OUT	: KOSTAL_AF2024_Core_Settings.T_MaxString_UTF8;
	_resp	: KOSTAL_AF2024_Core_Settings.T_MaxString_UTF8;
	_split: KOSTAL_AF2024_Core_StringTools.FB_Split_UTF8;
	_udi: UDINT;
END_VAR

//cameras with InSigtVisionSuite sends MAC ID with ':'

_IN:= IN;

Tc2_Utilities.FindAndDeleteChar(ADR(_IN), '$0A', ADR(_resp), SIZEOF(_resp));
	
_split.Split_Delimiter(_resp, ':');

_OUT:= '';

FOR _udi:= _split.Results.NumberOfLines - 5 TO _split.Results.NumberOfLines DO

	_OUT:= Tc2_Standard.CONCAT(_OUT,  _split.Results.line_GET(_udi));

	IF _udi < _split.Results.NumberOfLines THEN	_OUT:= Tc2_Standard.CONCAT(_OUT,  ':');	END_IF

END_FOR

Tc2_Utilities.FindAndDeleteChar(ADR(_OUT), ' ', ADR(_resp), SIZEOF(_resp));

_catchMacId:= _resp;
END_METHOD

METHOD PROTECTED _getCommand : KOSTAL_AF2024_Core_Settings.T_MaxString_UTF8

VAR_INPUT
	ID				: E_Command_TcpIp;
	Parameter : KOSTAL_AF2024_Core_Settings.T_MaxString_UTF8;
END_VAR
VAR
	_c	: KOSTAL_AF2024_Core_StringTools.FB_Concat_UTF8;
END_VAR

IF ID = E_Command_TcpIp.GetFormatstring	THEN	
	_c.Clear();
	_c.addContent('GV');
	_c.addContent(_sheetName);
	_c.addContent('.A0$R$N');
	_getCommand:= _c.getResult();		//get formatted result(s)
//	_getCommand:= 'GVAF_2024.A0$R$N';		//get formatted result(s)
ELSE																				
	_getCommand:= SUPER^._getCommand(ID, Parameter);	
END_IF
END_METHOD

PROPERTY PUBLIC SheetName : KOSTAL_AF2024_Core_Settings.T_MaxString_UTF8
GET
SheetName := _sheetName;
END_GET
SET
_sheetName := SheetName;
END_SET
END_PROPERTY

END_FUNCTION_BLOCK
